{attribute 'analysis' := '-33'}
VAR_GLOBAL CONSTANT
    iSLAVEADDR_ARR_SIZE	: UINT := 256;
    ESC_MAX_PORTS : UINT := 3; // Maximum number of ports (4) on ESC
END_VAR

(* stored: Version 1.1.0.1
   GVL Global_Variables_EtherCAT: Id {d76f2eaf-f0c3-42c2-8317-22c7ba689cf7} *)
